// TIA Portal V20 export
Screen "RobotService_Zone01_2"  1276x673
  ScreenItem "Line_Header_X0_Y64" at 0,64 size 1280x0  Type=HmiLine
  ScreenItem "permanentareaborderrectangle" at 0,0 size 0x0  Type=HmiRectangle
  ScreenItem "Button_Back" at 2,2 size 90x60  Type=HmiButton
  ScreenItem "Title_ScreenOverview_X390_Y2_3" at 368,5 size 510x57  Type=HmiTextBox
  ScreenItem "120RB01" at 272,81 size 193x297  Type=HmiFaceplateContainer
  ScreenItem "160RB02" at 47,81 size 193x297  Type=HmiFaceplateContainer
  ScreenItem "Faceplate container_1" at 1127,70 size 127x580  Type=HmiFaceplateContainer
